// TIA Portal V20 export
// export: Created 2026-11-12T11:17:34.1461208Z, ExportSetting WithDefaults, DisplayName Totally Integrated Automation Portal, DisplayVersion V20, DisplayName TIA Portal Openness, DisplayVersion V20, DisplayName TIA Portal Teamcenter Gateway, DisplayVersion V20, DisplayName TIA Portal Version Control Interface, DisplayVersion V20, DisplayName STEP 7 Professional, DisplayVersion V20, DisplayName STEP 7 CFC, DisplayVersion V20, DisplayName STEP 7 Safety, DisplayVersion V20, DisplayName WinCC Basic/Comfort/Advanced, DisplayVersion V20, DisplayName SIMATIC Visualization Architect, DisplayVersion V20, DisplayName WinCC Professional, DisplayVersion V20, DisplayName SIMATIC Visualization Architect, DisplayVersion V20, DisplayName WinCC Unified, DisplayVersion V20, DisplayName SIMATIC Visualization Architect, DisplayVersion V20
TYPE "UDT_Entradas_RFID"
// stored: IsFailsafeCompliant false
   STRUCT
      Tag_datos_escritos : Bool;   // Datos escritos
      Tag_datos_leidos : Bool;   // Datos leidos
      Reservado_E4_2 : Bool;
      Reservado_E4_3 : Bool;
      Tag_antena_apagada : Bool;   // Antena apagada
      Tag_detectado : Bool;   // Tag detectado
      Tag_error : Bool;   // Error
      Tag_proceso_listo : Bool;   // Proceso listo
      Tag_codigo_error : Byte;   // Codigo de error
      Tag_direccion_confirmada : Word;   // Direccion de escritura
      Tag_datos_leidos_escritos : Array[0..27] of Byte;   // Datos
   END_STRUCT;
END_TYPE
